(* IEC 61131-3 sources: repolevel_ST_code_completion/dataset/project_code/Robotics_DynamicModel/struct, 2 files *)

(* ---- TwistVec.st ---- *)
/// A six dimensional twist vector representing
/// a generalized velocity or acceleration.
TYPE TwistVec :
STRUCT
    /// The angular velocity or acceleration component.
    w : SM3M.SMC_VECTOR3D;
    /// The linear velocity or acceleration component.
    v : SM3M.SMC_VECTOR3D;
END_STRUCT
END_TYPE

(* ---- WrendchVec.st ---- *)
/// A six dimensional wrench vector representing
/// a generalized momentum or force.
TYPE WrenchVec :
STRUCT
    /// The angular momentum or torque component.
    m : SM3M.SMC_VECTOR3D;
    /// The linear momentum or force component.
    f : SM3M.SMC_VECTOR3D;
END_STRUCT
END_TYPE
